FUNCTION_BLOCK SC_TemplateUntil (* TEMPLATE for the contract of your primitive, SC_<Primitive>: copy it under that name, then change what says YOUR OWN, and this comment; keep the rest as it is. The contract of a skill primitive, the only part that is its own: which command it sends (and with what argument, and which when it ends), how long it may run, and three conditions on the equipment's signals and its parameters: when it may start, when it is done, what must hold while it runs. Technical: TemplateUntil: Precondition TRUE; Template.MyCommand until MyInput; Invariant TRUE *)
  (* Standard: 61499-2 *)
  (* Version 0.1, 2026-09-28, Project contributors, AAU Smart Production Lab *)
  PACKAGE capping;
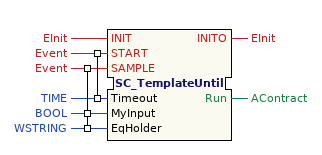
  EVENT_INPUT
    INIT : EInit; (* Initialise: name the OPC UA variables of the parameters and results *)
    START WITH Timeout; (* A run starts, with the parameters: say what the skill does *)
    SAMPLE WITH MyInput, EqHolder; (* The equipment's newest state arrived *)
  END_EVENT
  EVENT_OUTPUT
    INITO : EInit; (* Initialised: the next block of the INIT chain goes on *)
  END_EVENT
  VAR_INPUT
    Timeout : TIME; (* How long the run may take before it fails with Timeout (3) *)
    MyInput : BOOL; (* YOUR OWN, one per input pin. Template: MyInput, an input *)
    EqHolder : WSTRING; (* Who holds the equipment now (empty: free), passed on to the run *)
  END_VAR
  PLUGS
    Run : modlib::AContract; (* To the run (AContract): what the skill does and when it is done *)
  END_PLUGS
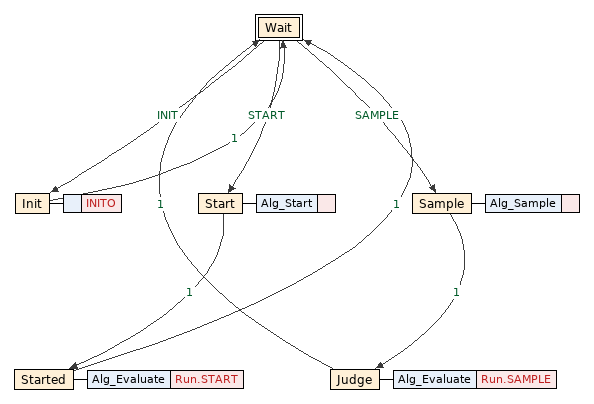
  EC_STATES
    Wait;
    Init : -> INITO;
    Start : Alg_Start;
    Started : Alg_Evaluate -> Run.START;
    Sample : Alg_Sample;
    Judge : Alg_Evaluate -> Run.SAMPLE;
  END_STATES
  EC_TRANSITIONS
    Wait TO Init := INIT;
    Init TO Wait := 1;
    Wait TO Start := START;
    Start TO Started := 1;
    Started TO Wait := 1;
    Wait TO Sample := SAMPLE;
    Sample TO Judge := 1;
    Judge TO Wait := 1;
  END_TRANSITIONS
  ALGORITHM Alg_Start IN ST:
Run.Timed := FALSE;  (* YOUR OWN: TRUE: the time RunTime ends the run; FALSE: Run.Post ends it, and RunTime is its timeout *)
Run.RunTime := Timeout;  (* YOUR OWN: how long it runs (Timed) or may run (not Timed) *)
Run.Command := 1;  (* YOUR OWN: the command to send: its number in EC_, in the order of its table (0 Stop, 1 MyCommand, ...) *)
Run.Arg := 0.0;  (* YOUR OWN: the command's argument, e.g. a position; 0.0 for none *)
Run.StopCommand := 0;  (* YOUR OWN: the command sent when the run ends: 0 Stop (all off), or another *)
  END_ALGORITHM
  ALGORITHM Alg_Evaluate IN ST:
Run.Pre := TRUE;  (* YOUR OWN: the precondition: may it start? *)
Run.Post := MyInput;  (* YOUR OWN: the postcondition: is it done? *)
Run.Inv := TRUE;  (* YOUR OWN: the invariant: may it go on? *)
  END_ALGORITHM
  ALGORITHM Alg_Sample IN ST:
Run.EqHolder := EqHolder;
  END_ALGORITHM
END_FUNCTION_BLOCK
